(* IEC 61131-3 sources: model-first-plc-agent-ai/results/T1-W-13, 2 files *)

(* ---- a1_code.st ---- *)
FUNCTION_BLOCK ConveyorRuntime
VAR_INPUT
    sensor_a : BOOL;
    sensor_b : BOOL;
END_VAR
VAR_OUTPUT
    conveyor : BOOL := FALSE;
END_VAR
VAR
    x0 : BOOL := TRUE;
    x1 : BOOL := FALSE;
    t1 : BOOL;
    t2 : BOOL;
    conveyor_latch : RS;
END_VAR

t1 := x0 AND sensor_a AND NOT sensor_b;
t2 := x1 AND sensor_b;

conveyor_latch(S := t1, R1 := t2);

x1 := conveyor_latch.Q1;
x0 := NOT x1;

conveyor := x1;

END_FUNCTION_BLOCK

PROGRAM Main
VAR
    SensorA AT %IX100.0 : BOOL;
    SensorB AT %IX100.1 : BOOL;
    Conveyor AT %QX100.0 : BOOL;
END_VAR
VAR
    runtime_logic : ConveyorRuntime;
END_VAR

runtime_logic(
    sensor_a := SensorA,
    sensor_b := SensorB
);

Conveyor := runtime_logic.conveyor;

END_PROGRAM

(* ---- a2_code.st ---- *)
FUNCTION_BLOCK FB_ConveyorControl
VAR_INPUT
    sensor_a : BOOL;
    sensor_b : BOOL;
END_VAR
VAR_OUTPUT
    conveyor : BOOL;
END_VAR
VAR
    run_latch : RS;
END_VAR

run_latch(
    S := sensor_a AND NOT sensor_b,
    R1 := sensor_b
);
conveyor := run_latch.Q1;

END_FUNCTION_BLOCK

PROGRAM Main
VAR
    sensor_a AT %IX100.0 : BOOL;
    sensor_b AT %IX100.1 : BOOL;
    conveyor AT %QX100.0 : BOOL;
END_VAR
VAR
    controller : FB_ConveyorControl;
END_VAR

controller(
    sensor_a := sensor_a,
    sensor_b := sensor_b
);
conveyor := controller.conveyor;

END_PROGRAM
